(* IEC 61131-3 sources: plcassist-cli/packages/volt-lsp-iec/test-corpus/lenze-mid/Device/Plc Logic/Application/Library Manager/L_SEMP_ErrorManagement, 29 files *)

(* ---- L_SEMP_EVENTIDS.gvl ---- *)
VAR_GLOBAL
	CMPID_CMPLENZEERRORMANAGEMENTACCESS : DWORD := 16#2014;
	EVT_CMPLENZEERRORMANAGEMENTACCESSACTSTATEDETERMINEEVENTCHANGED : DWORD := 16#10000011;
	EVTPARAMID_CMPLENZEERRORMANAGEMENTACCESSACTSTATEDETERMINEEVENTCHANGED : WORD := 16#1;
	EVTVERSION_CMPLENZEERRORMANAGEMENTACCESSACTSTATEDETERMINEEVENTCHANGED : WORD := 16#1;
	EVT_CMPLENZEERRORMANAGEMENTACCESSRESETOCCURRED : DWORD := 16#10000012;
	EVTPARAMID_CMPLENZEERRORMANAGEMENTACCESSRESETOCCURRED : WORD := 16#1;
	EVTVERSION_CMPLENZEERRORMANAGEMENTACCESSRESETOCCURRED : WORD := 16#1;
	EVT_CMPLENZEERRORMANAGEMENTACCESSCOMMANDEVENTREACTION : DWORD := 16#10000013;
	EVTPARAMID_CMPLENZEERRORMANAGEMENTACCESSCOMMANDEVENTREACTION : WORD := 16#1;
	EVTVERSION_CMPLENZEERRORMANAGEMENTACCESSCOMMANDEVENTREACTION : WORD := 16#1;
	EVT_CMPLENZEERRORMANAGEMENTACCESSREADACTERRORDATAAVAILABLE : DWORD := 16#10000014;
	EVTPARAMID_CMPLENZEERRORMANAGEMENTACCESSREADACTERRORDATAAVAILABLE : WORD := 16#1;
	EVTVERSION_CMPLENZEERRORMANAGEMENTACCESSREADACTERRORDATAAVAILABLE : WORD := 16#1;
END_VAR

(* ---- GETBOOLEANPROPERTY.fun ---- *)
FUNCTION GETBOOLEANPROPERTY : BOOL
VAR_INPUT
	STKEY : WSTRING;
END_VAR
END_FUNCTION

(* ---- GETCOMPANY.fun ---- *)
FUNCTION GETCOMPANY : WSTRING
END_FUNCTION

(* ---- GETNUMBERPROPERTY.fun ---- *)
FUNCTION GETNUMBERPROPERTY : DINT
VAR_INPUT
	STKEY : WSTRING;
END_VAR
END_FUNCTION

(* ---- GETTEXTPROPERTY.fun ---- *)
FUNCTION GETTEXTPROPERTY : WSTRING
VAR_INPUT
	STKEY : WSTRING;
END_VAR
END_FUNCTION

(* ---- GETTEXTPROPERTY2.fun ---- *)
FUNCTION GETTEXTPROPERTY2 : POINTER TO WSTRING
VAR_INPUT
	STKEY : WSTRING;
END_VAR
END_FUNCTION

(* ---- GETTITLE.fun ---- *)
FUNCTION GETTITLE : WSTRING
END_FUNCTION

(* ---- GETVERSION.fun ---- *)
FUNCTION GETVERSION : VERSION
END_FUNCTION

(* ---- GETVERSIONPROPERTY.fun ---- *)
FUNCTION GETVERSIONPROPERTY : VERSION
VAR_INPUT
	STKEY : WSTRING;
END_VAR
END_FUNCTION

(* ---- L_SEMP_CLEAREVENT.fun ---- *)
FUNCTION L_SEMP_CLEAREVENT : RTS_IEC_RESULT
VAR_INPUT
	HHANDLE : RTS_IEC_HANDLE := RTS_INVALID_HANDLE;
	UIEVENTID : UINT := 16#0;
END_VAR
END_FUNCTION

(* ---- L_SEMP_CLEAREVENT_V2.fun ---- *)
FUNCTION L_SEMP_CLEAREVENT_V2 : RTS_IEC_RESULT
VAR_INPUT
	HHANDLE : RTS_IEC_HANDLE := RTS_INVALID_HANDLE;
	UIEVENTID : UINT := 16#0;
	UITEXTREFID : UINT := 16#0;
END_VAR
END_FUNCTION

(* ---- L_SEMP_GETACCESSACTSTATEDETERMINEPARAMETER.fun ---- *)
FUNCTION L_SEMP_GETACCESSACTSTATEDETERMINEPARAMETER : BOOL
VAR_INPUT
	PPARAMETER : POINTER TO BYTE;
	SEVERITY : POINTER TO USINT;
	EVENTID : POINTER TO WORD;
	TEXTREFID : POINTER TO WORD;
	ACTSTATEDETERMINEEVENT : POINTER TO DWORD;
END_VAR
END_FUNCTION

(* ---- L_SEMP_GETACCESSACTSTATEDETERMINEPARAMETER2.fun ---- *)
FUNCTION L_SEMP_GETACCESSACTSTATEDETERMINEPARAMETER2 : BOOL
VAR_INPUT
	PPARAMETER : POINTER TO BYTE;
	SEVERITY : POINTER TO USINT;
	EVENTID : POINTER TO WORD;
	TEXTREFID : POINTER TO WORD;
	ACTSTATEDETERMINEEVENT : POINTER TO DWORD;
	ACTERRORCODE : POINTER TO DWORD;
END_VAR
END_FUNCTION

(* ---- L_SEMP_GETACCESSACTSTATEDETERMINEPARAMETER3.fun ---- *)
FUNCTION L_SEMP_GETACCESSACTSTATEDETERMINEPARAMETER3 : BOOL
VAR_INPUT
	PPARAMETER : POINTER TO BYTE;
	SEVERITY : POINTER TO USINT;
	EVENTID : POINTER TO WORD;
	TEXTREFID : POINTER TO WORD;
	ACTSTATEDETERMINEEVENT : POINTER TO DWORD;
	ACTERRORCODE : POINTER TO DWORD;
	USERGROUP : POINTER TO USINT;
END_VAR
END_FUNCTION

(* ---- L_SEMP_GETCOMMANDEVENTREACTIONPARAMETER.fun ---- *)
FUNCTION L_SEMP_GETCOMMANDEVENTREACTIONPARAMETER : BOOL
VAR_INPUT
	PPARAMETER : POINTER TO BYTE;
	SEVERITY : POINTER TO USINT;
	EVENTID : POINTER TO WORD;
	TEXTREFID : POINTER TO WORD;
END_VAR
END_FUNCTION

(* ---- L_SEMP_GETRESETOCUREDINCOMPONENT.fun ---- *)
FUNCTION L_SEMP_GETRESETOCUREDINCOMPONENT : BOOL
VAR_INPUT
	PPARAMETER : POINTER TO BYTE;
	PCOMPONENT : POINTER TO DWORD;
	PACTSEVERITY : POINTER TO USINT;
END_VAR
END_FUNCTION

(* ---- L_SEMP_NOTIFYEVENT.fun ---- *)
FUNCTION L_SEMP_NOTIFYEVENT : RTS_IEC_RESULT
VAR_INPUT
	HHANDLE : RTS_IEC_HANDLE := RTS_INVALID_HANDLE;
	UIEVENTID : UINT := 16#0;
	ESEVERITY : L_SEMP_Serverity := L_SEMP_Serverity.LEM_SEV_NO_RESPONSE;
	UITEXTREFID : UINT := 16#0;
	UINUMPARAM : UINT := 16#0;
	PPARAMETES : POINTER TO L_SEMP_EventParameters;
END_VAR
END_FUNCTION

(* ---- L_SEMP_NOTIFYEVENT_V2.fun ---- *)
FUNCTION L_SEMP_NOTIFYEVENT_V2 : RTS_IEC_RESULT
VAR_INPUT
	HHANDLE : RTS_IEC_HANDLE := RTS_INVALID_HANDLE;
	UIEVENTID : UINT := 16#0;
	ESEVERITY : USINT := L_SEMP_Serverity.LEM_SEV_NO_RESPONSE;
	UITEXTREFID : UINT := 16#0;
	UINUMPARAM : UINT := 16#0;
	PPARAMETES : POINTER TO L_SEMP_EventParameters;
	UIEVENTCONTROL : UINT := 16#0;
	UIUSERPRIORITY : UINT := 16#0;
	UITARGETGROUP : UINT := 16#0;
END_VAR
END_FUNCTION

(* ---- L_SEMP_NOTIFYEVENTSHORT.fun ---- *)
FUNCTION L_SEMP_NOTIFYEVENTSHORT : RTS_IEC_RESULT
VAR_INPUT
	HHANDLE : RTS_IEC_HANDLE := RTS_INVALID_HANDLE;
	UIEVENTID : UINT := 16#0;
	ESEVERITY : L_SEMP_Serverity := L_SEMP_Serverity.LEM_SEV_NO_RESPONSE;
	UITEXTREFID : UINT := 16#0;
	UINUMPARAM : UINT := 16#0;
	PPARAMETES : POINTER TO L_SEMP_EventParametersShort;
END_VAR
END_FUNCTION

(* ---- L_SEMP_NOTIFYEVENTSHORT_V2.fun ---- *)
FUNCTION L_SEMP_NOTIFYEVENTSHORT_V2 : RTS_IEC_RESULT
VAR_INPUT
	HHANDLE : RTS_IEC_HANDLE := RTS_INVALID_HANDLE;
	UIEVENTID : UINT := 16#0;
	ESEVERITY : L_SEMP_Serverity := L_SEMP_Serverity.LEM_SEV_NO_RESPONSE;
	UITEXTREFID : UINT := 16#0;
	UINUMPARAM : UINT := 16#0;
	PPARAMETES : POINTER TO L_SEMP_EventParametersShort;
	UIEVENTCONTROL : UINT := 16#0;
	UIUSERPRIORITY : UINT;
	UITARGETGROUP : UINT := 16#0;
END_VAR
END_FUNCTION

(* ---- L_SEMP_NOTIFYEVENTSHORT_V3.fun ---- *)
FUNCTION L_SEMP_NOTIFYEVENTSHORT_V3 : RTS_IEC_RESULT
VAR_INPUT
	HHANDLE : RTS_IEC_HANDLE := RTS_INVALID_HANDLE;
	UIEVENTID : UINT := 16#0;
	ESEVERITY : L_SEMP_Serverity := L_SEMP_Serverity.LEM_SEV_NO_RESPONSE;
	UITEXTREFID : UINT := 16#0;
	UINUMPARAM : UINT := 16#0;
	PPARAMETES : POINTER TO L_SEMP_EventParametersShort;
	UIEVENTCONTROL : UINT := 16#0;
	UIREACTION : UINT := 0;
	UITARGETGROUP : UINT := 16#0;
END_VAR
END_FUNCTION

(* ---- L_SEMP_REGISTERCOMPONENT.fun ---- *)
FUNCTION L_SEMP_REGISTERCOMPONENT : RTS_IEC_HANDLE
VAR_INPUT
	SCOMPONENTNAME : STRING := '';
	UILAYER : UINT := 16#0;
	UITEXTREFID : UINT := 16#0;
	UIREAKTIONITF : UINT := 16#0;
END_VAR
END_FUNCTION

(* ---- L_SEMP_REGISTERCOMPONENT2.fun ---- *)
FUNCTION L_SEMP_REGISTERCOMPONENT2 : RTS_IEC_HANDLE
VAR_INPUT
	SCOMPONENTNAME : STRING := '';
	UILAYER : UINT := 16#0;
	UITEXTREFID : UINT := 16#0;
	UIREAKTIONITF : UINT := 16#0;
	UIGETALLRESETS : UINT := 16#0;
END_VAR
END_FUNCTION

(* ---- L_SEMP_REQUESTRESET.fun ---- *)
FUNCTION L_SEMP_REQUESTRESET : RTS_IEC_RESULT
VAR_INPUT
	HHANDLE : RTS_IEC_HANDLE := RTS_INVALID_HANDLE;
END_VAR
END_FUNCTION

(* ---- L_SEMP_REQUESTRESETCOMPONENT.fun ---- *)
FUNCTION L_SEMP_REQUESTRESETCOMPONENT : RTS_IEC_RESULT
VAR_INPUT
	HHANDLE : RTS_IEC_HANDLE := RTS_INVALID_HANDLE;
END_VAR
END_FUNCTION

(* ---- L_SEMP_REQUESTRESETCOMPONENTLIST.fun ---- *)
FUNCTION L_SEMP_REQUESTRESETCOMPONENTLIST : RTS_IEC_RESULT
VAR_INPUT
	HANDLELIST : POINTER TO RTS_IEC_HANDLE;
	LISTCOUNT : WORD;
END_VAR
END_FUNCTION

(* ---- L_SEMP_UNREGISTERCOMPONENT.fun ---- *)
FUNCTION L_SEMP_UNREGISTERCOMPONENT : RTS_IEC_RESULT
VAR_INPUT
	HHANDLE : RTS_IEC_HANDLE := RTS_INVALID_HANDLE;
END_VAR
END_FUNCTION

(* ---- L_SEMP_READACTUALERRORCODE.fb ---- *)
FUNCTION_BLOCK L_SEMP_READACTUALERRORCODE
VAR_INPUT
	XENABLE : BOOL;
END_VAR
VAR_OUTPUT
	XBUSY : BOOL;
	DWERRORCODE : DWORD;
	ESEVERITY : L_SEMP_ServerityLevel;
END_VAR
VAR
	ITFCALLBACK : CmpEventMgr.ICmpEventCallback;
	HEVENTUPDATEACTIVEERROR : RTS_IEC_HANDLE := SysTypes.RTS_INVALID_HANDLE;
	HINTERFACEUPDATEACTIVEERROR : RTS_IEC_HANDLE := SysTypes.RTS_INVALID_HANDLE;
	WEVTCOUNT_UPDATEACTIVEERROR : WORD;
	SEVERITY_INT : USINT;
	EVENTID_INT : WORD;
	USERGROUP_INT : USINT;
	EUSERGROUP : USINT;
	TEXTREFID_INT : WORD;
	ACTSTATEDETERMINEEVENT_INT : DWORD;
	ACTERRORCODE_INT : DWORD;
	USERGROUP : USINT;
END_VAR
END_FUNCTION_BLOCK

METHOD FB_EXIT : BOOL
VAR_INPUT
	BINCOPYCODE : BOOL;
END_VAR
END_METHOD

METHOD FB_INIT : BOOL
VAR_INPUT
	BINITRETAINS : BOOL;
	BINCOPYCODE : BOOL;
END_VAR
END_METHOD

METHOD EVENTCALLBACK : UDINT
VAR_INPUT
	PEVENTPARAM : POINTER TO EventParam;
END_VAR
END_METHOD

METHOD REGISTEREVENT
END_METHOD

METHOD UNREGISTEREVENT
END_METHOD

(* ---- L_SEMP_SETERROR.fb ---- *)
FUNCTION_BLOCK L_SEMP_SETERROR
VAR_INPUT
	XRESETERROR : BOOL;
	XSETERROR1 : BOOL;
	ESEVERITY1 : L_SEMP_ServerityLevel;
	WERRORID1 : WORD;
	WTEXTREFID1 : WORD;
	XSETERROR2 : BOOL;
	ESEVERITY2 : L_SEMP_ServerityLevel;
	WERRORID2 : WORD;
	WTEXTREFID2 : WORD;
	XSETERROR3 : BOOL;
	ESEVERITY3 : L_SEMP_ServerityLevel;
	WERRORID3 : WORD;
	WTEXTREFID3 : WORD;
	XSETERROR4 : BOOL;
	ESEVERITY4 : L_SEMP_ServerityLevel;
	WERRORID4 : WORD;
	WTEXTREFID4 : WORD;
END_VAR
VAR_OUTPUT
	XERROR : BOOL;
	EERRORID : L_IE1P_Error;
	XERRORRESETACTIVE : BOOL;
END_VAR
VAR
	ERRORHANDLE : RTS_IEC_HANDLE := 0;
	ELAYER : L_SEMP_Layer := L_SEMP_Layer.Application;
	EERRORBEHAVIOUR : L_SEMP_Behaviour := L_SEMP_Behaviour.ProcessErrorReaction;
	SCOMPONENTNAME : STRING := '';
	WDEFAULTTEXTREFID : WORD := 16#2C00;
	XDEFAULTTEXTREFIDVALID : BOOL;
	XRESETERROROLD : BOOL;
	XSETERROR1OLD : BOOL;
	XSETERROR2OLD : BOOL;
	XSETERROR3OLD : BOOL;
	XSETERROR4OLD : BOOL;
	SINSTANCESTR : STRING;
	SINSTANCESTRDUMMY : STRING;
	ESEVERITY1_INT : L_SEMP_ServerityLevel;
	ESEVERITY2_INT : L_SEMP_ServerityLevel;
	ESEVERITY3_INT : L_SEMP_ServerityLevel;
	ESEVERITY4_INT : L_SEMP_ServerityLevel;
	WERRORID1_INT : WORD;
	WERRORID2_INT : WORD;
	WERRORID3_INT : WORD;
	WERRORID4_INT : WORD;
	ITFCALLBACK : CmpEventMgr.ICmpEventCallback;
	HEVENTRESETOCCURED : RTS_IEC_HANDLE := SysTypes.RTS_INVALID_HANDLE;
	HINTERFACERESETOCCURED : RTS_IEC_HANDLE := SysTypes.RTS_INVALID_HANDLE;
	WEVTCOUNT_RESETOCCURED : WORD;
	XRESETOCCURED : BOOL;
	XFBERRORINT1 : BOOL;
	EFBERRORIDINT1 : L_IE1P_Error;
	XFBERRORINT2 : BOOL;
	EFBERRORIDINT2 : L_IE1P_Error;
	XFBERRORINT3 : BOOL;
	EFBERRORIDINT3 : L_IE1P_Error;
	XFBERRORINT4 : BOOL;
	EFBERRORIDINT4 : L_IE1P_Error;
	COMPONENTNAME : STRING;
	DEFAULTTEXTREFID : WORD;
	ERRORBEHAVIOUR : L_SEMP_Behaviour;
	LAYER : L_SEMP_Layer;
END_VAR
END_FUNCTION_BLOCK

METHOD CHECKSETERROR : STRING
VAR_IN_OUT
	XSETERROR : BOOL;
	XSETERROROLD : BOOL;
	ESEVERITY : L_SEMP_Serverity;
	ESEVERITY_INT : L_SEMP_Serverity;
	WERRORID : WORD;
	WERRORID_INT : WORD;
	WTEXTREFID : WORD;
	XFBERRORINT : BOOL;
	EFBERRORIDINT : L_IE1P_Error;
END_VAR
END_METHOD

METHOD GETINSTANCENAME : STRING
END_METHOD

METHOD FB_AFTERINIT
END_METHOD

METHOD FB_EXIT : BOOL
VAR_INPUT
	BINCOPYCODE : BOOL;
END_VAR
END_METHOD

METHOD FB_INIT : BOOL
VAR_INPUT
	BINITRETAINS : BOOL;
	BINCOPYCODE : BOOL;
END_VAR
END_METHOD

METHOD EVENTCALLBACK : UDINT
VAR_INPUT
	PEVENTPARAM : POINTER TO EventParam;
END_VAR
END_METHOD

METHOD REGISTEREVENT
END_METHOD

METHOD UNREGISTEREVENT
END_METHOD
